(* IEC 61131-3 sources: genai_codesys/experiments/raw/formal/20261109_234635_2ba96d/public_01/codex_cli__deepseek-v4.1-flash-1017/attempt_00, 2 files *)

(* ---- declaration.st ---- *)
FUNCTION_BLOCK FB_AutomatedFillingLine
VAR_INPUT
    bottleSensor : BOOL;
    cleaningConfirmButton : BOOL;
    fillingConfirmButton : BOOL;
    cappingConfirmButton : BOOL;
    packingConfirmButton : BOOL;
    finishedButton : BOOL;
END_VAR
VAR_OUTPUT
    Pump_Motor : BOOL;
    Filling_Valve : BOOL;
    Capping_Machine : BOOL;
    Packing_Machine : BOOL;
    Completion_Light : BOOL;
END_VAR
VAR
    iState : INT := 0;
END_VAR
END_FUNCTION_BLOCK

(* ---- implementation.st ---- *)
CASE iState OF
    0:
        IF bottleSensor THEN
            iState := 1;
        END_IF;
    1:
        IF cleaningConfirmButton THEN
            iState := 2;
        END_IF;
    2:
        IF fillingConfirmButton THEN
            iState := 3;
        END_IF;
    3:
        IF cappingConfirmButton THEN
            iState := 4;
        END_IF;
    4:
        IF packingConfirmButton THEN
            iState := 5;
        END_IF;
    5:
        IF finishedButton THEN
            iState := 0;
        END_IF;
END_CASE

Pump_Motor := (iState = 1);
Filling_Valve := (iState = 2);
Capping_Machine := (iState = 3);
Packing_Machine := (iState = 4);
Completion_Light := (iState = 5);
